(* IEC 61131-3 sources: 2026_Projet_YGO_ExcavatriceDragage/CODE_BACKUP/CODE_20260822_IntroductionTestCI/D_JOYSTICK, 4 files *)

(* ---- ST_Joystick_AxisCmd.st ---- *)
(* =======================================================================
   🕹️ ST_Joystick_AxisCmd — Consigne d'axe normalisée (sortie FB_Joystick)
   ───────────────────────────────────────────────────────────────
   🎯 Rôle : Structure de consigne d'axe 4 champs produite par FB_Joystick.
   📤 Champs : Enable, StartStop, SpeedRef, Direction.
   📄 Doc métier : DOC/AF/AF_Partie-08_Fonction_Joystick_v2.0.md
   ======================================================================= *)

TYPE ST_Joystick_AxisCmd :
STRUCT
    // === CONSIGNES DE PILOTAGE AXE ===
    Enable      : BOOL;   // --> [CMD] Autorisation globale pipeline (FALSE=neutralisation, sorties coupees)
    StartStop   : BOOL;   // --> [CMD] Validation de mouvement (TRUE=acceleration, FALSE=deceleration)
    SpeedRef    : REAL;   // --> [CMD] Consigne vitesse signee (-100.0..+100.0 %, signe coherent avec Direction)
    Direction   : INT;    // --> [CMD] Sens de mouvement (-1=Arriere/Descente, 0=Neutre, +1=Avant/Montee)
END_STRUCT
END_TYPE

(* ---- FB_AxisScale.st ---- *)
(* =======================================================================
   ⚙️ FB_AxisScale — Normalisation et zone morte d'un axe joystick
   ───────────────────────────────────────────────────────────────
   🎯 Rôle : Normalise une valeur brute (0..10000) selon le neutre calibré
             et applique une zone morte en unités brutes (compte ADC).
   🛡️ Garde-fou : Saturation stricte de la consigne à +/-100.0 %.
   📄 Doc métier : DOC/AF/AF_Partie-08_Fonction_Joystick_v2.0.md
   ======================================================================= *)

FUNCTION_BLOCK FB_AxisScale
VAR_INPUT
    // === ENTRÉES MESURÉES & CONFIGURATION ===
    RawIn       : INT;  // --> [HW]  Valeur brute potentiometre/Hall (0..10000)
    Neutral     : INT;  // --> [CFG] Point milieu calibre (compte brut ADC)
    DeadbandRaw : INT;  // --> [CFG] Zone morte en unites brutes ADC (ex: 300)
END_VAR
VAR_OUTPUT
    // === CONSIGNES CALCULÉES ===
    OutPct      : REAL; // <-- [STAT] Consigne d'axe mise a l'echelle (-100.0..+100.0 %)
END_VAR
VAR
    // === VARIABLES LOCALES INTERNES ===
    Delta       : REAL; // . [LOC]  Amplitude utile de la demi-plage d'axe
END_VAR

IF RawIn >= Neutral THEN
    Delta := INT_TO_REAL(10000 - Neutral);
    IF Delta > 0.0 THEN
        OutPct := (INT_TO_REAL(RawIn - Neutral) / Delta) * 100.0;
    ELSE
        OutPct := 0.0;
    END_IF;
ELSE
    Delta := INT_TO_REAL(Neutral);
    IF Delta > 0.0 THEN
        OutPct := (INT_TO_REAL(RawIn - Neutral) / Delta) * 100.0;
    ELSE
        OutPct := 0.0;
    END_IF;
END_IF;

IF ABS(RawIn - Neutral) <= DeadbandRaw THEN
    OutPct := 0.0;
END_IF;

// 🛡️ Limitation de plage : une valeur brute hors plage nominale ne doit jamais
// produire une consigne supérieure à ±100 %. Ce garde-fou protège les
// consommateurs en aval, notamment la translation M3.
OutPct := LIMIT(-100.0, OutPct, 100.0);

(* ---- FB_Filter_PT1.st ---- *)
(* =======================================================================
   ⚙️ FB_Filter_PT1 — Filtre passe-bas premier ordre (PT1 numérique)
   ───────────────────────────────────────────────────────────────
   🎯 Rôle : Filtre exponentiel discret y[k] = a*x[k] + (1-a)*y[k-1]
             avec a = CycleTimeS / (T + CycleTimeS). Pass-through si T=0 ou Cycle=0.
   📄 Doc métier : DOC/AF/AF_Partie-08_Fonction_Joystick_v2.0.md
   ======================================================================= *)

FUNCTION_BLOCK FB_Filter_PT1
VAR_INPUT
    // === CONSIGNES DE PILOTAGE & CONFIGURATION ===
    ValueIn    : REAL;  // --> [CMD] Consigne d'axe brute a filtrer
    TimeConst  : TIME;  // --> [CFG] Constante de temps du filtre (ex: T#200ms)
    CycleTimeS : REAL;  // --> [CFG] Temps de cycle reel de la tache en secondes (ex: 0.02)
END_VAR
VAR_OUTPUT
    // === SORTIES LISSÉES ===
    ValueOut   : REAL;  // <-- [STAT] Consigne d'axe lissee par filtre PT1
END_VAR
VAR
    // === VARIABLES LOCALES INTERNES ===
    T          : REAL;  // . [LOC]  Constante de temps convertie en secondes
    Alpha      : REAL;  // . [LOC]  Facteur d'attenuation du filtre exponentiel
END_VAR

T := TIME_TO_REAL(TimeConst) / 1000.0; // ms → s

IF T <= 0.0 OR CycleTimeS <= 0.0 THEN
    ValueOut := ValueIn;
ELSE
    Alpha    := CycleTimeS / (T + CycleTimeS);
    ValueOut := Alpha * ValueIn + (1.0 - Alpha) * ValueOut;
END_IF;

(* ---- FB_Joystick.st ---- *)
(* =======================================================================
   🕹️ FB_Joystick — Acquisition & conditionnement du geste opérateur
   ───────────────────────────────────────────────────────────────
   🎯 Rôle : Acquisition 2 axes Hall + bouton homme-mort normatif.
             Pipeline par axe : FB_AxisScale -> FB_Filter_PT1 -> Homme-Mort -> ST_Joystick_AxisCmd.
   🔒 Sécurité : Armement homme-mort par maintien au neutre.
                 Désarmement sur neutre prolongé, changement mode ou fin benne.
   📤 Sorties : AxisCmdX/Y, signaux de diagnostic et miroirs maintenance.
   📄 Doc métier : DOC/AF/AF_Partie-08_Fonction_Joystick_v2.0.md
   ======================================================================= *)

FUNCTION_BLOCK FB_Joystick
VAR_INPUT
    // === PERMIS SÉCURITÉ & ETATS SYSTEME ===
    Enable                    : BOOL;       // --> [CMD]  Active la logique du bloc (TRUE=Autorise)
    Reset                     : BOOL;       // --> [CMD]  Acquittement defaut
    PowerContactorEngaged     : BOOL;       // --> [SAFE] Conditions globales OK (chaine AU rearmee)
    Mode                      : E_Mode;     // --> [SAFE] Changement de mode desarme l'homme-mort
    BenneBusy                 : BOOL;       // --> [SAFE] Fin de cycle benne (front descendant) desarme l'homme-mort
    PreserveArmingAfterBucket : BOOL;       // --> [SAFE] Maintien armement pendant fermeture ExtractionSequence

    // === ACQUISITION MATERIELLE & DIAGNOSTIC ===
    BusCanOpenOP              : ST_Diag_Device; // --> [HW]   Etat presence noeud CAN
    JoystickOP                : ST_Diag_Device; // --> [HW]   Mode esclave CANopen actif
    RawX                      : INT;        // --> [HW]   Valeur brute axe X (0..10000)
    RawY                      : INT;        // --> [HW]   Valeur brute axe Y (0..10000)
    RawButton                 : BOOL;       // --> [HW]   Etat brut bouton homme-mort

    // === COMMANDES OPÉRATEUR & CALIBRATION ===
    BtnCalibrate              : BOOL;       // --> [CMD]  Demande de recalage neutre

    // === REGLAGES & CONFIGURATION ===
    InvertX                   : BOOL := FALSE;   // --> [CFG]  Inversion sens de l'axe X
    InvertY                   : BOOL := FALSE;   // --> [CFG]  Inversion sens de l'axe Y
    DeadbandRaw               : INT := 300;      // --> [CFG]  Zone morte en points ADC bruts (0..10000)
    FilterTime                : TIME := T#0MS;   // --> [CFG]  Filtrage premier ordre axe
    NeutralHoldTime           : TIME := T#100MS; // --> [CFG]  Maintien continu au neutre avant desarmement
    DeadmanArmHoldTime        : TIME := T#100MS; // --> [CFG]  Appui continu bouton requis pour armer
    DeadmanArmGraceTime       : TIME := T#3S;    // --> [CFG]  Delai de grace post-armement avant desarmement neutre
END_VAR
VAR_OUTPUT
    // === ETATS IEC & SYNOPTIQUE ===
    Ready                     : BOOL;       // <-- [STAT] FB pret a fonctionner
    Busy                      : BOOL;       // <-- [STAT] Traitement en cours
    Done                      : BOOL;       // <-- [STAT] Donnees valides disponibles
    Button                    : BOOL;       // <-- [STAT] Bouton homme-mort filtre

    // === DIAGNOSTIC & ANOMALIES ===
    Error                     : BOOL;       // <-- [DIAG] Presence anomalie
    ErrorId                   : WORD;       // <-- [DIAG] Bit0: Echec calibration Joystick (RawX/Y hors plage)

    // === CONSIGNES AXES NORMALISEES ===
    AxisCmdX                  : ST_Joystick_AxisCmd; // <-- [ACT]  Sortie normalisee axe X
    AxisCmdY                  : ST_Joystick_AxisCmd; // <-- [ACT]  Sortie normalisee axe Y

    // === MESURES & MIROIRS MAINTENANCE ===
    NeutralXAct               : INT;        // <-- [STAT] Point neutre X actuel pour IHM/Test
    NeutralYAct               : INT;        // <-- [STAT] Point neutre Y actuel pour IHM/Test
    SpeedXPct                 : REAL;       // <-- [STAT] Consigne vitesse axe X signee (-100..+100 %), miroir AxisCmdX.SpeedRef
    DirectionX                : INT;        // <-- [STAT] Sens axe X (-1=Rev/0=Neutre/+1=Fwd), miroir AxisCmdX.Direction
    SpeedYPct                 : REAL;       // <-- [STAT] Consigne vitesse axe Y signee (-100..+100 %), miroir AxisCmdY.SpeedRef
    DirectionY                : INT;        // <-- [STAT] Sens axe Y (-1=Rev/0=Neutre/+1=Fwd), miroir AxisCmdY.Direction
    DeadmanArmed              : BOOL;       // <-- [STAT] Geste arme (bouton appuye au neutre) - IHM/diagnostic
    AtNeutral                 : BOOL;       // <-- [STAT] TRUE si les 2 axes sont en zone morte (position centrale)
END_VAR
VAR_IN_OUT
    // === RETENTION & CALIBRATION PERSISTANTE ===
    NeutralXMem               : INT;        // <-> [BUS]  Point neutre X persistant global
    NeutralYMem               : INT;        // <-> [BUS]  Point neutre Y persistant global
END_VAR
VAR
    // === SOUS-INSTANCES FB & TIMERS ===
    CycleTimeCalc             : FB_CycleTime;        // * [INST] Calcul du temps de cycle reel
    ScaleX                    : FB_AxisScale;        // * [INST] Normalisation et zone morte axe X
    ScaleY                    : FB_AxisScale;        // * [INST] Normalisation et zone morte axe Y
    FilterX                   : FB_Filter_PT1;       // * [INST] Filtre passe-bas PT1 axe X
    FilterY                   : FB_Filter_PT1;       // * [INST] Filtre passe-bas PT1 axe Y
    ResetEdge                 : R_TRIG;              // * [INST] Detecteur front montant Reset
    DeadmanEdge               : R_TRIG;              // * [INST] Detecteur front montant Bouton homme-mort
    NeutralHoldTimer          : TON;                 // * [INST] Temporisation maintien au neutre
    DeadmanArmTimer           : TON;                 // * [INST] Temporisation maintien bouton armement
    DeadmanArmGraceTimer      : TON;                 // * [INST] Temporisation delai de grace post-armement
    BenneBusyFallEdge         : F_TRIG;              // * [INST] Detecteur front descendant Fin de cycle benne

    // === VARIABLES LOCALES INTERNES ===
    CmdXVal                   : REAL;                // . [LOC]  Consigne axe X calculee apres filtrage/homme-mort
    CmdYVal                   : REAL;                // . [LOC]  Consigne axe Y calculee apres filtrage/homme-mort
    LastCalibrate             : BOOL;                // . [LOC]  Memorisation etat precedent bouton calibration
    DeadmanArmPending         : BOOL;                // . [LOC]  Armement en cours d'attente de la tempo maintien
    LastMode                  : E_Mode;              // . [LOC]  Memorisation mode scan precedent pour detection changement
END_VAR

{region "§1 Gate securite"}
// 🛑 1. GATE (Sécurités et coupures prioritaires)
IF NOT Enable OR NOT PowerContactorEngaged OR NOT BusCanOpenOP.Operational OR NOT JoystickOP.Operational THEN
    Ready := FALSE; Busy := FALSE; Done := FALSE;
    AxisCmdX.Enable := FALSE; AxisCmdX.StartStop := FALSE; AxisCmdX.SpeedRef := 0.0; AxisCmdX.Direction := 0;
    AxisCmdY.Enable := FALSE; AxisCmdY.StartStop := FALSE; AxisCmdY.SpeedRef := 0.0; AxisCmdY.Direction := 0;
    SpeedXPct := 0.0; DirectionX := 0;
    SpeedYPct := 0.0; DirectionY := 0;
    Button := FALSE;
    AtNeutral := TRUE;
    DeadmanArmed := FALSE;
    DeadmanArmPending := FALSE;
    NeutralHoldTimer(IN := FALSE, PT := NeutralHoldTime);
    DeadmanArmTimer(IN := FALSE, PT := DeadmanArmHoldTime);
    DeadmanArmGraceTimer(IN := FALSE, PT := DeadmanArmGraceTime);
    NeutralXAct := NeutralXMem;
    NeutralYAct := NeutralYMem;
    LastMode := Mode;   // Pas de faux changement détecté à la réactivation
    RETURN;
END_IF;

Ready := TRUE; Busy := TRUE;

{endregion}

{region "§2 Reset acquisition timing et bouton"}
// 🔑 2. RESET DÉFAUT (front + cause disparue, Partie3 §5)
ResetEdge(CLK := Reset);
IF ResetEdge.Q AND (RawX >= 2000 AND RawX <= 8000 AND RawY >= 2000 AND RawY <= 8000) THEN
    ErrorId := ErrorId AND 16#FFFE;
END_IF;

// 📥 3. ACQUISITION TIMING & BOUTON
CycleTimeCalc();
Button := RawButton;

{endregion}

{region "§3 Calibration et mise a echelle"}
// 🎯 4. CALIBRATION DYNAMIQUE (Zone RETAIN)
IF BtnCalibrate AND NOT LastCalibrate THEN
    IF RawX >= 2000 AND RawX <= 8000 AND RawY >= 2000 AND RawY <= 8000 THEN
        NeutralXMem := RawX;
        NeutralYMem := RawY;
    ELSE
        // Un seul bit pour une seule cause (Partie3 §3)
        ErrorId := ErrorId OR 16#0001;
    END_IF;
END_IF;
Error := (ErrorId <> 16#0000);
LastCalibrate := BtnCalibrate;

// 🧮 4bis. MISE À L'ÉCHELLE (avant homme-mort — le neutre s'évalue sur les 2 axes déjà deadbandés)
ScaleX(RawIn := RawX, Neutral := NeutralXMem, DeadbandRaw := DeadbandRaw);
ScaleY(RawIn := RawY, Neutral := NeutralYMem, DeadbandRaw := DeadbandRaw);
AtNeutral := (ScaleX.OutPct = 0.0) AND (ScaleY.OutPct = 0.0);   // IHM/diagnostic — position centrale (zone morte)

{endregion}

{region "§4 Desarmements changement mode et fin benne"}
// 4ter-bis. CHANGEMENT DE MODE : désarme le homme-mort dès que Mode change
// (MAINT_N1/N2/SEMI_AUTO/AUTO). Évite qu'une commande en cours traverse le changement
// de mode et soit réinterprétée soudainement. Repassage par le neutre + nouvel appui exigé.
IF Mode <> LastMode THEN
    DeadmanArmed := FALSE;
    DeadmanArmPending := FALSE;   // Nouvel appui exigé après changement de mode
END_IF;
LastMode := Mode;

// 4ter-ter. FIN DE CYCLE BENNE : désarmement général pour qu'une fermeture manuelle
// ne démarre jamais M1/M2 par surprise. Exception : ExtractionSequence garde l'armement
// pendant sa fermeture (enchaînement palier 1 sous ses propres interlocks synchro/position).
BenneBusyFallEdge(CLK := BenneBusy);
IF BenneBusyFallEdge.Q AND NOT PreserveArmingAfterBucket THEN
    DeadmanArmed := FALSE;
    DeadmanArmPending := FALSE;   // Nouvel appui exigé après fin de cycle benne
END_IF;

{endregion}

{region "§5 Armement homme mort"}
// 4ter. BOUTON HOMME-MORT — armement par MAINTIEN (DeadmanArmHoldTime), indépendant de la
// position des axes pendant l'appui.
// Armement par MAINTIEN (DeadmanArmHoldTime), indépendant de la position des axes pendant
// l'appui : appui (front) → maintien 100 ms → armé, quelle que soit la position des axes durant
// ce maintien. Relâchement AVANT la fin du maintien = tentative annulée (DeadmanArmPending
// retombe), un nouvel appui (front) est requis — pas d'armement différé "surprise" sur un appui
// prolongé après un désarmement (mode/benne/neutre). Sûr même si le joystick est déjà hors zone
// morte à la fin du maintien : les rampes d'accel/décel restent gérées par les FB aval
// (FB_Winch/FB_Translation), donc pas de démarrage brutal possible côté ce FB.
DeadmanEdge(CLK := RawButton);
IF DeadmanEdge.Q THEN
    DeadmanArmPending := TRUE;
END_IF;
IF NOT RawButton THEN
    DeadmanArmPending := FALSE;
END_IF;

// 🛡️ SÉCURITÉ C4 (ISO 13849) : armement STRICTEMENT conditionné par DeadmanArmPending.
// Tout désarmement (changement de mode, fin de cycle benne, passage neutre prolongé)
// efface DeadmanArmPending et EXIGE un nouvel appui conscient (front montant de RawButton).
DeadmanArmTimer(IN := DeadmanArmPending AND NOT DeadmanArmed, PT := DeadmanArmHoldTime);
IF DeadmanArmTimer.Q THEN
    DeadmanArmed := TRUE;
    DeadmanArmPending := FALSE;
END_IF;

// ⏱️ 4bis. GESTION DU DÉSARMEMENT PAR MAINTIEN AU NEUTRE
DeadmanArmGraceTimer(IN := DeadmanArmed, PT := DeadmanArmGraceTime);
NeutralHoldTimer(IN := DeadmanArmed AND AtNeutral AND DeadmanArmGraceTimer.Q,
                 PT := NeutralHoldTime);
IF NeutralHoldTimer.Q THEN
    DeadmanArmed := FALSE;      // Neutre maintenu après la grâce = désarmement
END_IF;

{endregion}

{region "§6 Pipeline axe X"}
// 🕹️ 5. PIPELINE TRAITEMENT — AXE X
IF InvertX THEN
    FilterX(ValueIn := -ScaleX.OutPct, TimeConst := FilterTime, CycleTimeS := CycleTimeCalc.CycleTimeS);
ELSE
    FilterX(ValueIn := ScaleX.OutPct, TimeConst := FilterTime, CycleTimeS := CycleTimeCalc.CycleTimeS);
END_IF;

// Consigne forcée à 0.0 tant que le geste n'est pas armé (homme-mort)
CmdXVal := SEL(DeadmanArmed, 0.0, FilterX.ValueOut);

// Mapping Sortie Standardisée Axe X
AxisCmdX.Enable := TRUE;
AxisCmdX.SpeedRef := CmdXVal;
AxisCmdX.StartStop := (ABS(CmdXVal) > 0.1);

IF CmdXVal > 0.1 THEN
    AxisCmdX.Direction := 1;
ELSIF CmdXVal < -0.1 THEN
    AxisCmdX.Direction := -1;
ELSE
    AxisCmdX.Direction := 0;
    AxisCmdX.SpeedRef := 0.0;
END_IF;

// Miroirs maintenance
SpeedXPct := AxisCmdX.SpeedRef;
DirectionX := AxisCmdX.Direction;

{endregion}

{region "§7 Pipeline axe Y et sorties"}
// 🕹️ 6. PIPELINE TRAITEMENT — AXE Y
IF InvertY THEN
    FilterY(ValueIn := -ScaleY.OutPct, TimeConst := FilterTime, CycleTimeS := CycleTimeCalc.CycleTimeS);
ELSE
    FilterY(ValueIn := ScaleY.OutPct, TimeConst := FilterTime, CycleTimeS := CycleTimeCalc.CycleTimeS);
END_IF;

// Consigne forcée à 0.0 tant que le geste n'est pas armé (homme-mort)
CmdYVal := SEL(DeadmanArmed, 0.0, FilterY.ValueOut);

// Mapping Sortie Standardisée Axe Y
AxisCmdY.Enable := TRUE;
AxisCmdY.SpeedRef := CmdYVal;
AxisCmdY.StartStop := (ABS(CmdYVal) > 0.1);

IF CmdYVal > 0.1 THEN
    AxisCmdY.Direction := 1;
ELSIF CmdYVal < -0.1 THEN
    AxisCmdY.Direction := -1;
ELSE
    AxisCmdY.Direction := 0;
    AxisCmdY.SpeedRef := 0.0;
END_IF;

// Miroirs maintenance
SpeedYPct := AxisCmdY.SpeedRef;
DirectionY := AxisCmdY.Direction;

// 📤 7. VALIDATION DES SORTIES ÉTAT
NeutralXAct := NeutralXMem;
NeutralYAct := NeutralYMem;
Done := NOT Error;

{endregion}
